// TIA Portal project "Study-Project" (V14)

(* hardware
DEVICE "S71500/ET200MP station_1"  S7-1500 station
   slot 0: "Rail_0"  Rack  6ES7 590-1***0-0AA0
   slot 1: "PLC_1"  CPU 1511-1 PN  6ES7 511-1AK01-0AB0  V2.1
      slot 3: "CPU display_1"  6ES7591-1AA00-0AA0
   slot 2: "DI 16x24VDC HF_1"  DI 16x24VDC HF  6ES7 521-1BH00-0AB0  V2.1
   slot 3: "DQ 16x24VDC/0.5A ST_1"  DQ 16x24VDC/0.5A ST  6ES7 522-1BH00-0AB0  V2.0
   slot 4: "AI 4xU/I/RTD/TC ST_1"  AI 4xU/I/RTD/TC ST  6ES7 531-7QD00-0AB0  V1.0
   slot 5: "AQ 2xU/I ST_1"  AQ 2xU/I ST  6ES7 532-5NB00-0AB0  V1.0
DEVICE "HMI_1"  KTP400F Mobile
   slot 0: "KTP400F Mobile"  KTP400F Mobile  6AV2 125-2DB23-0AX0  14.0.1.0
   slot 1: "HMI_RT_1"  KTP400F Mobile  6AV2 125-2DB23-0AX0  14.0.1.0
   slot 5: "HMI_1.IE_CP_1"  PROFINET Interface  14.0.1.0
      slot 1: "PROFINET Interface_1"  PROFINET Interface
         slot 1: "Port_1"  Port
DEVICE "PC station"  SIMATIC PC station
   slot 0: "PC station"  Rail  SIMATIC PC-Station  V1.0
      slot 125: "Stationmanager"  Station_Manager  V6.0.4
*)

// ===== PLC "PLC_1"  CPU 1511-1 PN =====

VAR_GLOBAL   // PLC tag table "Default tag table"
   "E_Stop" AT %I0.0 : Bool;   // Emergency stop, normally closed wiring. 1 = healthy, 0 = pressed or wire broken
   "Mode_Auto" AT %I0.1 : Bool;   // Mode selector. 1 = auto, 0 = manual
   "Start" AT %I0.2 : Bool;   // Start button, normally open. TRUE while pressed
   "Stop" AT %I0.3 : Bool;   // Stop button, normally open wiring. 0 = healthy
   "Reset" AT %I0.4 : Bool;   // Reset button. Combined with HMI_Reset into Reset_Req
   "IR_Prox" AT %I0.5 : Bool;   // Product sensor. Each rising edge counts one product
   "Conveyor_Motor" AT %Q0.0 : Bool;   // Motor output, driven by Network 4
   "Diverter_Solenoid" AT %Q0.1 : Bool;   // 1 = reject
   "Alarm_Beacon" AT %Q0.2 : Bool;   // Alarm lamp. Driven by Alarm_Active OR E_Stop_Latched
   "Buzzer" AT %Q0.3 : Bool;
   "Load_Cell" AT %IW64 : Int;   // Load cell raw count, 4-20 mA. 5530 = 4 mA, 27648 = 20 mA
   "Speed_Feedback" AT %IW66 : Int;   // 0–10 V
   "VFD_Speed_Cmd" AT %QW80 : Int;   // Speed command to VFD. 27648 = 10 V = full speed
   "Arm_Spare" AT %QW82 : Int;   // Unused
   "HMI_Start" AT %M0.0 : Bool;   // Screen Start button, pressed = 1
   "HMI_Stop" AT %M0.1 : Bool;   // Screen Stop button, pressed = 1
   "HMI_Reset" AT %M0.2 : Bool;   // Screen Reset button, pressed = 1
   "Reset_Req" AT %M0.3 : Bool;   // Combined reset from the physical and screen buttons
   "HMI_Weight" AT %MD10 : Real;   // Weight copy for the HMI display
   "HMI_Accepted" AT %MW20 : Int;   // Accepted count copy for the HMI display
   "HMI_Rejected" AT %MW22 : Int;   // Reject count copy for the HMI display
   "HMI_Batch" AT %MW24 : Int;   // Remaining batch count copy for the HMI display
   "HMI_Alarm" AT %M4.0 : Bool;   // Sorter alarm copy for the HMI display
   "HMI_Latch" AT %M4.1 : Bool;   // E-stop latch copy for the HMI display
   "HMI_Speed_Pct" AT %MW26 : Int;   // Speed command, percent of full scale
   "HMI_RejectPct" AT %MD30 : Real;
   "HMI_Throughput" AT %MD34 : Real;
END_VAR

DATA_BLOCK "DB_Configuration"   // DB1
{ S7_Optimized_Access := 'TRUE' }
VERSION : 0.1
   VAR
      Weight_Limit_kg : Real := 25.0;
      Ramp_Up_Time : Time := T#5s;
      E_Stop_Grace : Time := T#2s;
      Batch_Size : Int := 50;
      Speed_Setpoint : Int := 27648;
      Sim_Enable : Bool := FALSE;
      Sim_Gap : Time := T#3s;
      Sim_Dwell : Time := T#1s;
      Sim_Light_Raw : Int := 16000;
      Sim_Heavy_Raw : Int := 24000;
      Sim_Heavy_Every : Int := 3;
   END_VAR
BEGIN
END_DATA_BLOCK

DATA_BLOCK "DB_Runtime"   // DB2
{ S7_Optimized_Access := 'TRUE' }
VERSION : 0.1
   VAR
      E_Stop_Latched : Bool;
      Weight_kg : Real;
      Total_Count : DInt;
      Alarm_Log : Array[1..20] of String[40];
      Manual_Mode : Bool;
      Log_Index : Int := 1;
      Load_Fault_Prev : Bool := FALSE;
      Reject_Count : Int;
      Batch_Remaining : Int;
      Alarm_Active : Bool;
      Accepted_Count : Int;
      Speed_Fault_Prev : Bool := FALSE;
      Run_Min : Real;
      Calc_Status : Int;
   END_VAR
BEGIN
END_DATA_BLOCK

DATA_BLOCK "FB_ProductSimulator_DB"   // DB3
{ S7_Optimized_Access := 'TRUE' }
VERSION : 0.1
// stored: InstanceOfName FB_ProductSimulator
"FB_ProductSimulator"
BEGIN
END_DATA_BLOCK

DATA_BLOCK "FB_ConveyorController_DB"   // DB4
{ S7_Optimized_Access := 'TRUE' }
VERSION : 0.1
// stored: InstanceOfName FB_ConveyorController
"FB_ConveyorController"
BEGIN
END_DATA_BLOCK

DATA_BLOCK "FB_SorterLogic_DB_1"   // DB5
{ S7_Optimized_Access := 'TRUE' }
VERSION : 0.1
// stored: InstanceOfName FB_SorterLogic
"FB_SorterLogic"
BEGIN
END_DATA_BLOCK

FUNCTION_BLOCK "FB_ConveyorController"   // FB1, SCL
{ S7_Optimized_Access := 'TRUE' }
VERSION : 0.1
   VAR_INPUT
      Run_Enable : Bool;
      Mode_Auto : Bool;
      Weight_kg : Real;
      Speed_Setpoint_Raw : Int;
   END_VAR
   VAR_OUTPUT
      VFD_Speed_Cmd : Int;
      Mode_Changed : Bool;
      Ramp_Done : Bool;
   END_VAR
   VAR
      Ramp_Up : TON_TIME;
      Stop_Grace : TOF_TIME;
      Mode_Prev : Bool;
      State : Word := W#16#0001;
   END_VAR
   VAR_TEMP
      Load_Factor : Real;
      Fraction : Real;
      Target : Real;
   END_VAR
BEGIN
   // Ramp-up on start and stop grace on stop, both driven by the run command
   #Ramp_Up(IN := #Run_Enable,
            PT := "DB_Configuration".Ramp_Up_Time);
   #Stop_Grace(IN := #Run_Enable,
               PT := "DB_Configuration".E_Stop_Grace);

   // XOR flags a manual-to-auto or auto-to-manual change for one scan
   #Mode_Changed := #Mode_Auto XOR #Mode_Prev;
   #Mode_Prev := #Mode_Auto;

   // One-hot state ring: bit 0 stopped, bit 1 ramping, bit 2 running, bit 3 stopping
   // ROL moves the active bit to the next state
   IF #State = W#16#0001 AND #Run_Enable THEN
       #State := ROL(IN := #State, N := 1);
   ELSIF #State = W#16#0002 AND #Ramp_Up.Q THEN
       #State := ROL(IN := #State, N := 1);
   ELSIF #State = W#16#0002 AND NOT #Run_Enable THEN
       // A stop during ramp-up skips straight to the grace period
       #State := W#16#0008;
   ELSIF #State = W#16#0004 AND NOT #Run_Enable THEN
       #State := ROL(IN := #State, N := 1);
   ELSIF #State = W#16#0008 AND #Run_Enable THEN
       // A restart during the grace period resumes the ramp
       #State := W#16#0002;
   ELSIF #State = W#16#0008 AND NOT #Stop_Grace.Q THEN
       #State := W#16#0001;
   END_IF;

   // Fraction of full speed: rises during ramp-up, holds, falls during grace
   IF #State = W#16#0002 THEN
       #Fraction := DINT_TO_REAL(T_CONV(#Ramp_Up.ET)) / DINT_TO_REAL(T_CONV("DB_Configuration".Ramp_Up_Time));
   ELSIF #State = W#16#0004 THEN
       #Fraction := 1.0;
   ELSIF #State = W#16#0008 THEN
       #Fraction := 1.0 - DINT_TO_REAL(T_CONV(#Stop_Grace.ET)) / DINT_TO_REAL(T_CONV("DB_Configuration".E_Stop_Grace));
   ELSE
       #Fraction := 0.0;
   END_IF;
   #Fraction := LIMIT(MN := 0.0, IN := #Fraction, MX := 1.0);

   // MUL: the load factor drops to 0.5 as the weight reaches the limit
   #Load_Factor := 1.0 - 0.5 * (#Weight_kg / "DB_Configuration".Weight_Limit_kg);
   #Load_Factor := LIMIT(MN := 0.5, IN := #Load_Factor, MX := 1.0);

   // MUL: setpoint scaled by load and ramp fraction, written to the VFD
   #Target := INT_TO_REAL(#Speed_Setpoint_Raw) * #Load_Factor;
   #VFD_Speed_Cmd := REAL_TO_INT(#Target * #Fraction);

   #Ramp_Done := (#State = W#16#0004);
END_FUNCTION_BLOCK

FUNCTION_BLOCK "FB_SorterLogic"   // FB2, SCL
{ S7_Optimized_Access := 'TRUE' }
VERSION : 0.1
   VAR_INPUT
      Weight_kg : Real;
      Load_Raw : Int;
      Product_Present : Bool;
      Reset_Cmd : Bool;
   END_VAR
   VAR_OUTPUT
      Reject_Cmd : Bool;
      Alarm_Active : Bool;
      Accepted_Count : Int;
      Reject_Count : Int;
      Batch_Remaining : Int;
      Total_Weight : Real := 0.0;
   END_VAR
   VAR
      Product_Edge : R_TRIG;
      Total_Ctr : CTU_INT;
   END_VAR
   VAR RETAIN
      Reject_Ctr : CTU_INT;
      Batch_Ctr : CTD_INT;
      Alarm_Latch : Bool := FALSE;
   END_VAR
   VAR_TEMP
      Overweight : Bool;
      Sensor_Fault : Bool;
      Reject_Req : Bool;
      Accept_Req : Bool;
      Interlock_OK : Bool;
      Alarm_Trigger : Bool;
   END_VAR
BEGIN
   // R_TRIG gives one pulse as each product reaches the sensor
   #Product_Edge(CLK := #Product_Present);

   // GT: the weight is above the limit when it exceeds Weight_Limit_kg
   #Overweight := #Weight_kg > "DB_Configuration".Weight_Limit_kg;

   // EQ: a raw count of 0 means the load cell wire is broken
   #Sensor_Fault := (#Load_Raw = 0);

   // AND: reject a present product that is overweight, accept one that is within the limit
   #Reject_Req := #Product_Present AND #Overweight;
   #Accept_Req := #Product_Present AND NOT #Overweight;

   // NAND: the diverter may act only when reject and accept are not both requested
   #Interlock_OK := NOT (#Reject_Req AND #Accept_Req);
   #Reject_Cmd := #Reject_Req AND #Interlock_OK;

   // CTU counts every product and every reject
   #Total_Ctr(CU := #Product_Edge.Q,
              R := #Reset_Cmd,
              PV := 32767);
   #Reject_Ctr(CU := #Reject_Cmd,
               R := #Reset_Cmd,
               PV := 32767);

   // CTD counts the batch down and reloads it when it reaches zero
   #Batch_Ctr(CD := #Product_Edge.Q,
              LD := #Reset_Cmd OR (#Batch_Ctr.CV <= 0),
              PV := "DB_Configuration".Batch_Size);

   // SUB: accepted products are the total minus the rejects
   #Accepted_Count := #Total_Ctr.CV - #Reject_Ctr.CV;
   #Reject_Count := #Reject_Ctr.CV;
   #Batch_Remaining := #Batch_Ctr.CV;

   // ADD: running total of product weight, cleared by Reset
   IF #Product_Edge.Q THEN
       #Total_Weight := #Total_Weight + #Weight_kg;
   END_IF;
   IF #Reset_Cmd THEN
       #Total_Weight := 0.0;
   END_IF;

   // OR: alarm on an overweight product or a sensor fault
   #Alarm_Trigger := #Reject_Req OR #Sensor_Fault;

   // Latch: Reset clears the alarm and takes priority over a new trigger
   IF #Reset_Cmd THEN
       #Alarm_Latch := FALSE;
   ELSIF #Alarm_Trigger THEN
       #Alarm_Latch := TRUE;
   END_IF;
   #Alarm_Active := #Alarm_Latch;
END_FUNCTION_BLOCK

FUNCTION_BLOCK "FB_ProductSimulator"   // FB3, SCL
{ S7_Optimized_Access := 'TRUE' }
VERSION : 0.1
   VAR_INPUT
      Enable : Bool;
      Real_IR : Bool;
      Real_Load : Int;
      Gap : Time;
      Dwell : Time;
      Light_Raw : Int;
      Heavy_Raw : Int;
      Heavy_Every : Int;
   END_VAR
   VAR_OUTPUT
      Present_Out : Bool;
      Load_Out : Int;
   END_VAR
   VAR
      Gap_T : TON_TIME;
      Dwell_T : TON_TIME;
      Presence : Bool;
      Prev_Present : Bool;
      Product_Count : Int;
   END_VAR
BEGIN
   // Timers run every scan so they reset cleanly when the simulation is switched off
   #Gap_T(IN := #Enable AND NOT #Presence,
          PT := #Gap);
   #Dwell_T(IN := #Enable AND #Presence,
            PT := #Dwell);

   // The gap ends by placing a product in front of the sensor, and the dwell ends by removing it
   IF NOT #Enable THEN
       #Presence := FALSE;
   END_IF;
   IF #Gap_T.Q THEN
       #Presence := TRUE;
   END_IF;
   IF #Dwell_T.Q THEN
       #Presence := FALSE;
   END_IF;

   // Count each rising edge of the presence signal, so the load pattern follows the product number
   IF #Presence AND NOT #Prev_Present THEN
       #Product_Count := #Product_Count + 1;
   END_IF;
   #Prev_Present := #Presence;

   // Simulated values when enabled, physical inputs passed through when disabled
   IF #Enable THEN
       #Present_Out := #Presence;
       IF #Heavy_Every > 0 AND (#Product_Count MOD #Heavy_Every = 0) THEN
           #Load_Out := #Heavy_Raw;
       ELSE
           #Load_Out := #Light_Raw;
       END_IF;
   ELSE
       #Present_Out := #Real_IR;
       #Load_Out := #Real_Load;
   END_IF;
END_FUNCTION_BLOCK

FUNCTION "FC_ScaleAnalogInput" : Void   // FC1, SCL
{ S7_Optimized_Access := 'TRUE' }
VERSION : 0.1
   VAR_INPUT
      AI_Raw : Int;
   END_VAR
   VAR_OUTPUT
      Weight_kg : Real;
   END_VAR
BEGIN
   // Counts below 5530 mean the loop is under 4 mA, so report zero and let diagnostics flag the fault
   IF #AI_Raw < 5530 THEN
       #Weight_kg := 0.0;
   ELSE
       #Weight_kg := INT_TO_REAL(#AI_Raw - 5530) / 22118.0 * 50.0;
   END_IF;
END_FUNCTION

FUNCTION "FC_CalculateStatistics" : Int   // FC2, SCL
{ S7_Optimized_Access := 'TRUE' }
VERSION : 0.1
   VAR_INPUT
      Reject_Count : Int;
      Total_Count : Int;
      Elapsed_Min : Real;
   END_VAR
   VAR_OUTPUT
      Reject_Rate_Pct : Real;
      Throughput_Per_Min : Real;
   END_VAR
BEGIN
   // A zero total or zero elapsed time would divide by zero, so return status 1 without calculating
   IF #Total_Count = 0 OR #Elapsed_Min <= 0.0 THEN
       #Reject_Rate_Pct := 0.0;
       #Throughput_Per_Min := 0.0;
       #FC_CalculateStatistics := 1;
       RETURN;
   END_IF;

   // Reject rate as a percentage of all products, and throughput as products per minute
   #Reject_Rate_Pct := INT_TO_REAL(#Reject_Count) / INT_TO_REAL(#Total_Count) * 100.0;
   #Throughput_Per_Min := INT_TO_REAL(#Total_Count) / #Elapsed_Min;

   // Status 0 means the results are valid
   #FC_CalculateStatistics := 0;
END_FUNCTION

ORGANIZATION_BLOCK "Main"   // OB1, LAD, ProgramCycle
TITLE = "Main Program Sweep (Cycle)"
{ S7_Optimized_Access := 'TRUE' }
VERSION : 0.1
   VAR_INPUT
      Initial_Call : Bool;   // Initial call of this OB
      Remanence : Bool;   // =True, if remanent data are available
   END_VAR
BEGIN
END_ORGANIZATION_BLOCK

ORGANIZATION_BLOCK "OB 30"   // OB30, LAD, CyclicInterrupt
{ S7_Optimized_Access := 'TRUE' }
VERSION : 0.1
   VAR_INPUT
      Initial_Call : Bool;   // Initial call of this OB
      Event_Count : Int;   // Events discarded
   END_VAR
BEGIN

REGION Network 1
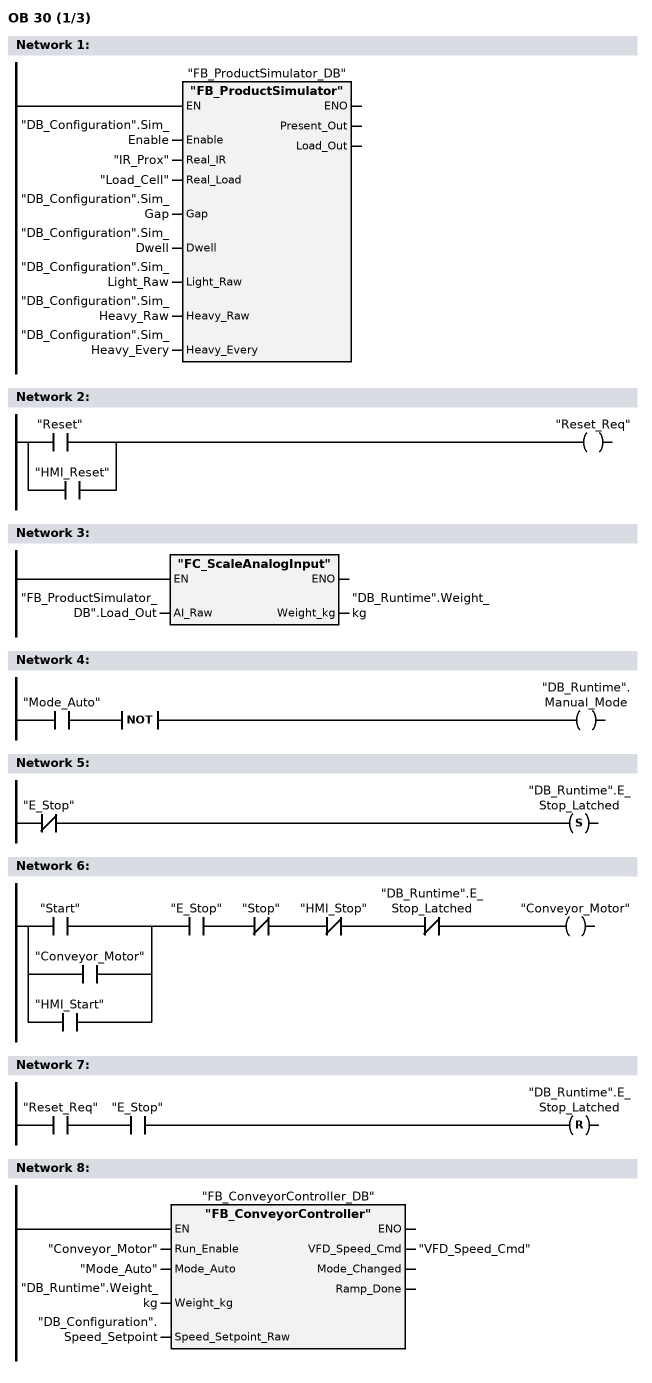
   RUNG wire#powerrail
      "FB_ProductSimulator_DB"(Enable := "DB_Configuration".Sim_Enable, Real_IR := "IR_Prox", Real_Load := "Load_Cell", Gap := "DB_Configuration".Sim_Gap, Dwell := "DB_Configuration".Sim_Dwell, Light_Raw := "DB_Configuration".Sim_Light_Raw, Heavy_Raw := "DB_Configuration".Sim_Heavy_Raw, Heavy_Every := "DB_Configuration".Sim_Heavy_Every, Present_Out =>, Load_Out =>)
   END_RUNG
   // the same network as SCL:
   "FB_ProductSimulator_DB"(Enable := "DB_Configuration".Sim_Enable,   // "FB_ProductSimulator"
                           Real_IR := "IR_Prox",
                           Real_Load := "Load_Cell",
                           Gap := "DB_Configuration".Sim_Gap,
                           Dwell := "DB_Configuration".Sim_Dwell,
                           Light_Raw := "DB_Configuration".Sim_Light_Raw,
                           Heavy_Raw := "DB_Configuration".Sim_Heavy_Raw,
                           Heavy_Every := "DB_Configuration".Sim_Heavy_Every);
END_REGION

REGION Network 2
   RUNG wire#powerrail
      Contact( "Reset" )
      wire#w1
      Coil( "Reset_Req" )
   END_RUNG
   RUNG wire#powerrail
      Contact( "HMI_Reset" )
   END_RUNG wire#w1
   // the same network as SCL:
   "Reset_Req" := "Reset" OR "HMI_Reset";
END_REGION

REGION Network 3
   RUNG wire#powerrail
      "FC_ScaleAnalogInput"(AI_Raw := "FB_ProductSimulator_DB".Load_Out, Weight_kg => "DB_Runtime".Weight_kg)
   END_RUNG
   // the same network as SCL:
   "FC_ScaleAnalogInput"(AI_Raw := "FB_ProductSimulator_DB".Load_Out, Weight_kg => "DB_Runtime".Weight_kg);
END_REGION

REGION Network 4
   RUNG wire#powerrail
      Contact( "Mode_Auto" )
      Not()
      Coil( "DB_Runtime".Manual_Mode )
   END_RUNG
   // the same network as SCL:
   "DB_Runtime".Manual_Mode := NOT "Mode_Auto";
END_REGION

REGION Network 5
   RUNG wire#powerrail
      I_Contact( "E_Stop" )
      S_Coil( "DB_Runtime".E_Stop_Latched )
   END_RUNG
   // the same network as SCL:
   IF NOT "E_Stop" THEN "DB_Runtime".E_Stop_Latched := TRUE; END_IF;
END_REGION

REGION Network 6
   RUNG wire#powerrail
      Contact( "Start" )
      wire#w1
      Contact( "E_Stop" )
      I_Contact( "Stop" )
      I_Contact( "HMI_Stop" )
      I_Contact( "DB_Runtime".E_Stop_Latched )
      Coil( "Conveyor_Motor" )
   END_RUNG
   RUNG wire#powerrail
      Contact( "Conveyor_Motor" )
   END_RUNG wire#w1
   RUNG wire#powerrail
      Contact( "HMI_Start" )
   END_RUNG wire#w1
   // the same network as SCL:
   "Conveyor_Motor" := ("Start" OR "Conveyor_Motor" OR "HMI_Start") AND "E_Stop" AND NOT "Stop" AND NOT "HMI_Stop" AND NOT "DB_Runtime".E_Stop_Latched;
END_REGION

REGION Network 7
   RUNG wire#powerrail
      Contact( "Reset_Req" )
      Contact( "E_Stop" )
      R_Coil( "DB_Runtime".E_Stop_Latched )
   END_RUNG
   // the same network as SCL:
   IF "Reset_Req" AND "E_Stop" THEN "DB_Runtime".E_Stop_Latched := FALSE; END_IF;
END_REGION

REGION Network 8
   RUNG wire#powerrail
      "FB_ConveyorController_DB"(Run_Enable := "Conveyor_Motor", Mode_Auto := "Mode_Auto", Weight_kg := "DB_Runtime".Weight_kg, Speed_Setpoint_Raw := "DB_Configuration".Speed_Setpoint, VFD_Speed_Cmd => "VFD_Speed_Cmd", Mode_Changed =>, Ramp_Done =>)
   END_RUNG
   // the same network as SCL:
   "FB_ConveyorController_DB"(Run_Enable := "Conveyor_Motor",   // "FB_ConveyorController"
                           Mode_Auto := "Mode_Auto",
                           Weight_kg := "DB_Runtime".Weight_kg,
                           Speed_Setpoint_Raw := "DB_Configuration".Speed_Setpoint,
                           VFD_Speed_Cmd => "VFD_Speed_Cmd");
END_REGION

REGION Network 9
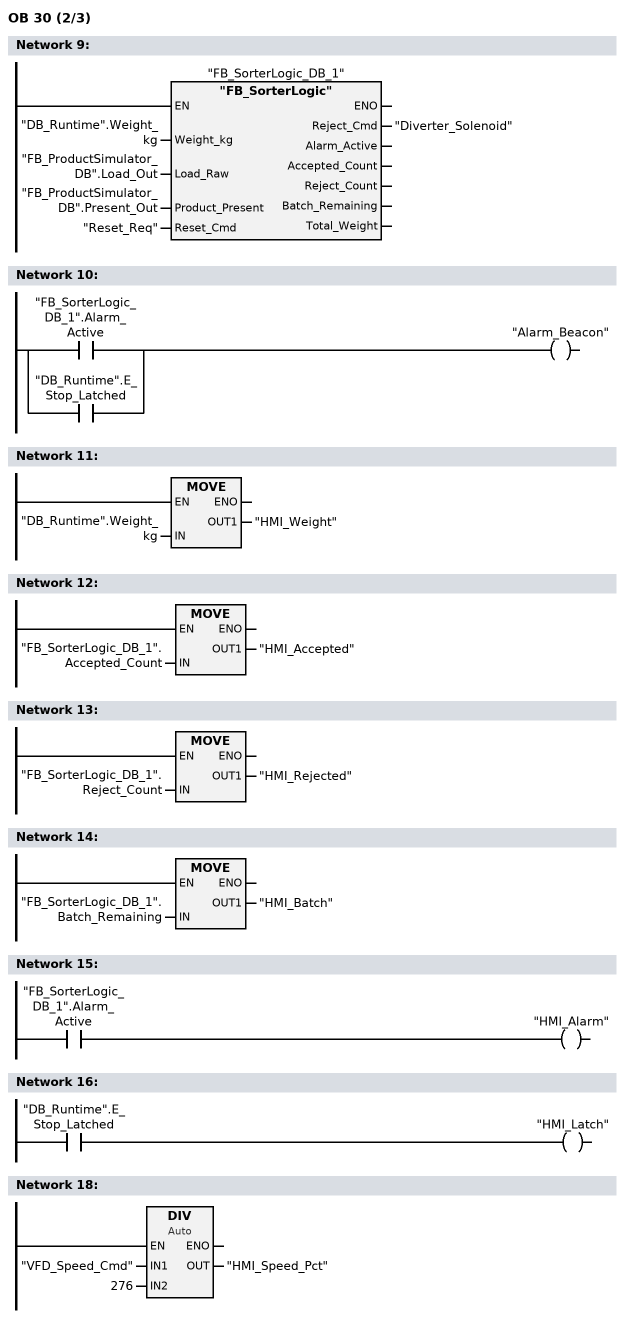
   RUNG wire#powerrail
      "FB_SorterLogic_DB_1"(Weight_kg := "DB_Runtime".Weight_kg, Load_Raw := "FB_ProductSimulator_DB".Load_Out, Product_Present := "FB_ProductSimulator_DB".Present_Out, Reset_Cmd := "Reset_Req", Reject_Cmd => "Diverter_Solenoid", Alarm_Active =>, Accepted_Count =>, Reject_Count =>, Batch_Remaining =>, Total_Weight =>)
   END_RUNG
   // the same network as SCL:
   "FB_SorterLogic_DB_1"(Weight_kg := "DB_Runtime".Weight_kg,   // "FB_SorterLogic"
                         Load_Raw := "FB_ProductSimulator_DB".Load_Out,
                         Product_Present := "FB_ProductSimulator_DB".Present_Out,
                         Reset_Cmd := "Reset_Req",
                         Reject_Cmd => "Diverter_Solenoid");
END_REGION

REGION Network 10
   RUNG wire#powerrail
      Contact( "FB_SorterLogic_DB_1".Alarm_Active )
      wire#w1
      Coil( "Alarm_Beacon" )
   END_RUNG
   RUNG wire#powerrail
      Contact( "DB_Runtime".E_Stop_Latched )
   END_RUNG wire#w1
   // the same network as SCL:
   "Alarm_Beacon" := "FB_SorterLogic_DB_1".Alarm_Active OR "DB_Runtime".E_Stop_Latched;
END_REGION

REGION Network 11
   RUNG wire#powerrail
      Move(in := "DB_Runtime".Weight_kg, out1 => "HMI_Weight")
   END_RUNG
   // the same network as SCL:
   "HMI_Weight" := "DB_Runtime".Weight_kg;
END_REGION

REGION Network 12
   RUNG wire#powerrail
      Move(in := "FB_SorterLogic_DB_1".Accepted_Count, out1 => "HMI_Accepted")
   END_RUNG
   // the same network as SCL:
   "HMI_Accepted" := "FB_SorterLogic_DB_1".Accepted_Count;
END_REGION

REGION Network 13
   RUNG wire#powerrail
      Move(in := "FB_SorterLogic_DB_1".Reject_Count, out1 => "HMI_Rejected")
   END_RUNG
   // the same network as SCL:
   "HMI_Rejected" := "FB_SorterLogic_DB_1".Reject_Count;
END_REGION

REGION Network 14
   RUNG wire#powerrail
      Move(in := "FB_SorterLogic_DB_1".Batch_Remaining, out1 => "HMI_Batch")
   END_RUNG
   // the same network as SCL:
   "HMI_Batch" := "FB_SorterLogic_DB_1".Batch_Remaining;
END_REGION

REGION Network 15
   RUNG wire#powerrail
      Contact( "FB_SorterLogic_DB_1".Alarm_Active )
      Coil( "HMI_Alarm" )
   END_RUNG
   // the same network as SCL:
   "HMI_Alarm" := "FB_SorterLogic_DB_1".Alarm_Active;
END_REGION

REGION Network 16
   RUNG wire#powerrail
      Contact( "DB_Runtime".E_Stop_Latched )
      Coil( "HMI_Latch" )
   END_RUNG
   // the same network as SCL:
   "HMI_Latch" := "DB_Runtime".E_Stop_Latched;
END_REGION

REGION Network 18
   RUNG wire#powerrail
      Div(in1 := "VFD_Speed_Cmd", in2 := 276, out => "HMI_Speed_Pct")
   END_RUNG
   // the same network as SCL:
   "HMI_Speed_Pct" := "VFD_Speed_Cmd" / 276;
END_REGION

REGION Network 19
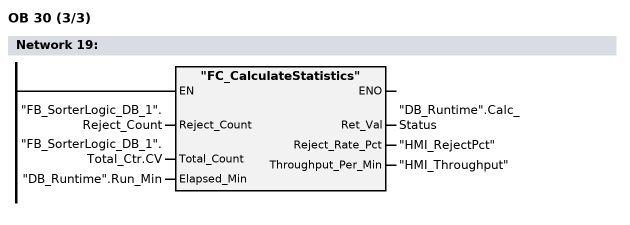
   RUNG wire#powerrail
      "FC_CalculateStatistics"(Reject_Count := "FB_SorterLogic_DB_1".Reject_Count, Total_Count := "FB_SorterLogic_DB_1".Total_Ctr.CV, Elapsed_Min := "DB_Runtime".Run_Min, Ret_Val => "DB_Runtime".Calc_Status, Reject_Rate_Pct => "HMI_RejectPct", Throughput_Per_Min => "HMI_Throughput")
   END_RUNG
   // the same network as SCL:
   "DB_Runtime".Calc_Status := "FC_CalculateStatistics"(Reject_Count := "FB_SorterLogic_DB_1".Reject_Count,
                           Total_Count := "FB_SorterLogic_DB_1".Total_Ctr.CV,
                           Elapsed_Min := "DB_Runtime".Run_Min,
                           Reject_Rate_Pct => "HMI_RejectPct",
                           Throughput_Per_Min => "HMI_Throughput");
END_REGION
END_ORGANIZATION_BLOCK

ORGANIZATION_BLOCK "Cyclic interrupt"   // OB35, SCL, CyclicInterrupt
{ S7_Optimized_Access := 'TRUE' }
VERSION : 0.1
   VAR_INPUT
      Initial_Call : Bool;   // Initial call of this OB
      Event_Count : Int;   // Events discarded
   END_VAR
   VAR_TEMP
      Load_Fault : Bool;
      Speed_Fault : Bool;
   END_VAR
BEGIN
   // Wire break: below 4 mA (5530 counts) means the loop is open
   #Load_Fault := "Load_Cell" < 5530;

   // Speed feedback must stay within 0 to 10 V (0 to 27648 counts)
   #Speed_Fault := "Speed_Feedback" < 0 OR "Speed_Feedback" > 27648;

   // Rising edge: the fault is present now and was absent on the previous run
   IF #Load_Fault AND NOT "DB_Runtime".Load_Fault_Prev THEN
       "DB_Runtime".Alarm_Log["DB_Runtime".Log_Index] := 'Load cell wire break';
       "DB_Runtime".Log_Index := "DB_Runtime".Log_Index + 1;
       IF "DB_Runtime".Log_Index > 20 THEN
           "DB_Runtime".Log_Index := 1;
       END_IF;
   END_IF;
   "DB_Runtime".Load_Fault_Prev := #Load_Fault;

   IF #Speed_Fault AND NOT "DB_Runtime".Speed_Fault_Prev THEN
       "DB_Runtime".Alarm_Log["DB_Runtime".Log_Index] := 'Speed feedback out of range';
       "DB_Runtime".Log_Index := "DB_Runtime".Log_Index + 1;
       IF "DB_Runtime".Log_Index > 20 THEN
           "DB_Runtime".Log_Index := 1;
       END_IF;
   END_IF;
   "DB_Runtime".Speed_Fault_Prev := #Speed_Fault;

   // Accumulate run time in minutes while the conveyor is running
   IF "Conveyor_Motor" THEN
       "DB_Runtime".Run_Min := "DB_Runtime".Run_Min + 5.0 / 60.0;
   END_IF;
END_ORGANIZATION_BLOCK

ORGANIZATION_BLOCK "Hardware interrupt"   // OB40, SCL, HWProcessInterruptExtended
{ S7_Optimized_Access := 'TRUE' }
VERSION : 0.1
   VAR_INPUT
      LADDR : Hw_Io;   // Hardware identifier
      USI : Word;   // User structure identifier
      IChannel : USInt;   // Interrupt channel number
      EventType : Byte;   // EventType
      PointAddr : DWord;
   END_VAR
BEGIN
   // Cut the motor immediately and latch the stop until Reset clears it
   "Conveyor_Motor" := FALSE;
   "DB_Runtime".E_Stop_Latched := TRUE;
END_ORGANIZATION_BLOCK

(* ===== HMI "HMI_RT_1" =====
system functions are stored by id; their names below are inferred from use
connection "HMI_Connection_1": ETHERNET, S7_1500_OMS

HMI tags "Default tag table"
   "Weight_kg" : Real = PLC HMI_Weight AT %MD10, 1 s
   "Tag_ScreenNumber_1" : UInt, internal
   "Speed_Pct" : Int = PLC HMI_Speed_Pct AT %MW26, 1 s
   "Accepted" : Int = PLC HMI_Accepted AT %MW20, 1 s
   "Rejected" : Int = PLC HMI_Rejected AT %MW22, 1 s
   "Batch_Left" : Int = PLC HMI_Batch AT %MW24, 1 s
   "Alarm" : Bool = PLC HMI_Alarm AT %M4.0, 1 s
   "Latch" : Bool = PLC HMI_Latch AT %M4.1, 1 s
   "Motor" : Bool = PLC Conveyor_Motor AT %Q0.0, 1 s
   "Btn_Start" : Bool = PLC HMI_Start AT %M0.0, 1 s
   "Btn_Stop" : Bool = PLC HMI_Stop AT %M0.1, 1 s
   "Btn_Reset" : Bool = PLC HMI_Reset AT %M0.2, 1 s
   "Reject_Pct" : Real = PLC HMI_RejectPct AT %MD30, 1 s
   "Throughput" : Real = PLC HMI_Throughput AT %MD34, 1 s

screen "Root screen" 480x231, template "Template_1"
   on GenerateScreen: SetTag("Weight_kg", 1)
   TextField "HmiScreenItemData" at 48,58 size 384x22; Text 'Welcome to HMI_1 (KTP400F Mobile)!'

Template "Template_1" 480x231
   Button "Exit" at 410,142 size 68x68; TextOff 'Exit'; PictureOff "ExitRuntime_KTP400F_Mobile_TR"; PictureOn "ExitRuntime_KTP400F_Mobile_TR"
      on Release: StopRuntime(0)
   Button "Template_Button" at 328,142 size 68x68; TextOff 'Text'
   Button "Template_Button_1" at 246,142 size 68x68; TextOff 'Text'
   Button "Template_Button_2" at 165,142 size 68x68; TextOff 'Text'
   Button "Alarms" at 83,142 size 68x68; TextOff 'Alarms'; PictureOff "AlarmDisplay_KTP400F_Mobile_TR"; PictureOn "AlarmDisplay_KTP400F_Mobile_TR"
      on Release: function_ef3f5d25("Alarm window_Unacknowledged", -1)
   Button "Start screen" at 1,142 size 68x68; TextOff 'Start screen'; PictureOff "NavigateHome_KTP400F_Mobile_TR"; PictureOn "NavigateHome_KTP400F_Mobile_TR"
      on Release: ActivateScreen("Root screen", 0)

screen "Dashboard" 480x231
   IOField "I/O field_1" at 112,9 size 96x32; FormatPattern 999
      ProcessValue <- "Weight_kg"
   TextField "Text field_1" at 12,15 size 93x20; Text 'Weight (kg)'
   IOField "I/O field_2" at 112,52 size 96x32; FormatPattern 99
      ProcessValue <- "Speed_Pct"
   TextField "Text field_2" at 12,58 size 84x20; Text 'Speed (%)'
   IOField "I/O field_3" at 112,96 size 96x32; FormatPattern 999
      ProcessValue <- "Accepted"
   TextField "Text field_3" at 12,102 size 75x20; Text 'Accepted'
   IOField "I/O field_4" at 112,139 size 96x32; FormatPattern 999
      ProcessValue <- "Rejected"
   TextField "Text field_4" at 12,145 size 71x20; Text 'Rejected'
   IOField "I/O field_5" at 365,12 size 96x32; FormatPattern 999
      ProcessValue <- "Batch_Left"
   TextField "Text field_5" at 265,18 size 82x20; Text 'Batch Left'
   IOField "I/O field_6" at 365,55 size 96x32; FormatPattern 99.99
      ProcessValue <- "Reject_Pct"
   TextField "Text field_9" at 265,61 size 87x20; Text 'Reject (%)'
   IOField "I/O field_7" at 365,99 size 96x32; FormatPattern 99.99
      ProcessValue <- "Throughput"
   TextField "Text field_11" at 265,99 size 96x36; Text 'Throughput (/min)'
   DateTimeField "Date/time field_1" at 259,140 size 202x29
   Button "Button_1" at 12,184 size 96x32; TextOff 'Start'
      on Release: ResetBit("Btn_Start")
      on Press: SetBit("Btn_Start")
   Button "Button_2" at 129,184 size 96x32; TextOff 'Stop'
      on Release: ResetBit("Btn_Stop")
      on Press: SetBit("Btn_Stop")
   Button "Button_3" at 247,184 size 96x32; TextOff 'Reset'
      on Release: ResetBit("Btn_Reset")
      on Press: SetBit("Btn_Reset")
   Button "Button_4" at 364,184 size 96x32; TextOff 'Menu'
*)